(* IEC 61131-3 sources: Testing02/Test_Version_Control/Temp/Import/TS_Test_UT/Logical/TS_UnitTest/Samples/Tests_Program/SPLMyCalc, 4 files *)

(* ---- SPLMyCalc.typ ---- *)
(********************************************************************
 * COPYRIGHT -- Bernecker + Rainer
 ********************************************************************
 * Library: SPLMyCalc
 * File: SPLMyCalc.typ
 * Author: B+R
 ********************************************************************
 * Data types of library SPLMyCalc
 ********************************************************************)

TYPE
	MyCalcOperator_enum :
		( (*Enumerator of maths operations*)
		splMyCalcOPERATOR_RESET_OUTPUTS := 0, (*Resets the outputs. No calculation*)
		splMyCalcOPERATOR_ADD := 1, (*Add *)
		splMyCalcOPERATOR_SUBTRACT := 2, (*Subtract*)
		splMyCalcOPERATOR_MULTIPLICATION := 3, (*Multiplication*)
		splMyCalcOPERATOR_DIVISION := 4, (*Division*)
		splMyCalcOPERATOR_SQUARE := 5, (*Square of Param 1*)
		splMyCalcOPERATOR_EXP := 6 (*Param1 ^ Param2*)
		);
END_TYPE

(* ---- SPLMyCalc.fun ---- *)
(********************************************************************
 * COPYRIGHT -- Bernecker + Rainer
 ********************************************************************
 * Library: SPLMyCalc
 * File: MyCalc.fun
 * Author: B+R
 ********************************************************************
 * Functions and function blocks of library SPLMyCalc
 ********************************************************************)

FUNCTION_BLOCK MyCalculator (*This functionblock provides several operations. If result is bigger / smaller than MIN or MAX, MIN or MAX are returned.*)
	VAR_INPUT
		CalcOperator : MyCalcOperator_enum; (*Calculation operation*)
		Param1 : INT; (*Paramerter 1*)
		Param2 : INT; (*Paramerter 2*)
	END_VAR
	VAR_OUTPUT
		Status : UINT; (*execution status: ERR_OK, ... *)
		Result : DINT; (*Result of the operation*)
	END_VAR
END_FUNCTION_BLOCK

(* ---- SPLMyCalc.st ---- *)
(********************************************************************
 * COPYRIGHT -- Bernecker + Rainer
 ********************************************************************
 * Library: SPLMyCalc
 * File: SPLMyCalc.st
 * Author: B+R
 ********************************************************************
 * Implementation of library SPLMyCalc
 ********************************************************************)

(* This can be used as a sample for  Test Driven Development (TDD)/ Test First Development
Steps (in a nutshell):
    o Define your API (FB, functions, ...)
		 this is already done for the FB MyCalc
	o Create a new test program (by using the template)
	o Write a test case (e.g. Addition) for this FB.
		The tests should describe the expected behavior.
	o Transfer the test program to the target and run the test in the test view
		The test case will fail
	o Implement this FB (Addition), build and transfer, then run the test again
		The test case will pass
	o Write next test (e.g. Subtraction).
	..
	o Write test for MIN / MAX (underflow/overflow)
   	o Run the tests to verify your implementation.

Note:
	The sample test program in SPL_MyCalcLib_C provides some test cases using this FB.

 *)
FUNCTION_BLOCK MyCalculator

	Status := ERR_NOTIMPLEMENTED;

END_FUNCTION_BLOCK

(* ---- SPLMyCalc.var ---- *)
(********************************************************************
 * COPYRIGHT --  Bernecker + Rainer
 ********************************************************************
 * Library: SPLMyCalc
 * File: SPLMyCalc.var
 * Author: B+R
 ********************************************************************
 * Constants of library SPLMyCalc
 ********************************************************************)
VAR CONSTANT
	splMyCalcERR_OUT_OF_RANGE : UINT := 50002;
	splMyCalcERR_NO_VALID_PARAM : UINT := 50001;
END_VAR
